Universal Robots PolyScope program: MainProg.urp

Program MainProg (createdIn=3.0.0 lastSavedIn=3.0.0 directory=/programs installation=default)
Robot Program (runOnlyOnce=true motionType=MoveJ speed=1.047198 acceleration=1.396263 useActiveTCP=false)
  'Program generated by VerticalBot Studio for UR10 on 25/10/2026 12:00:00'
  'Using nominal kinematics.'
  'Using Ref. Frame 2: p[-0.800000, 0.500000, 0.100000, 0.000000, 0.000000, 3.141593]'
  'Using TCP Paint gun: p[0.050000, 0.000000, 0.450000, 0.000000, 0.523599, 0.000000]'
  Script: set_tcp(p[0.050000, 0.000000, 0.450000, 0.000000, 0.523599, 0.000000])
  Call ApproachMove
  Call SprayOn
  Call PaintTop
  Call SprayOn
  Call Retract
SubProgram  [hidden by the author, left out]
SubProgram  [hidden by the author, left out]
SubProgram  [hidden by the author, left out]
SubProgram  [hidden by the author, left out]
SubProgram ApproachMove [hidden by the author, left out]
SubProgram SprayOn [hidden by the author, left out]
SubProgram PaintTop [hidden by the author, left out]
SubProgram Retract [hidden by the author, left out]
